(* IEC 61131-3 sources: trust-platform/examples/rust_barcode/src/generated, 1 file *)

(* ---- rust_pous.st ---- *)
(* GENERATED by trust-runtime from rust/src/lib.rs - do not edit *)
{attribute 'rust'}
FUNCTION_BLOCK GS1_LABEL
VAR_INPUT
    EN : BOOL := TRUE;
    code : STRING[64];
END_VAR
VAR_OUTPUT
    gtin : STRING[14];
    batch : STRING[20];
    expiry : DATE;
    gtin_ok : BOOL;
    error : INT;
    ENO : BOOL;
END_VAR
END_FUNCTION_BLOCK
